Fanuc KAREL source: KA00111.KL

PROGRAM KA00111
%NOLOCKGROUP
VAR
  SRC: CONFIG
  DST: BOOLEAN
BEGIN
  SRC.CFG_FLIP = TRUE
  DST = SRC
END KA00111
